SUBAPPLICATION Button_IXA_OR_AX_TO_DataPanel_QXA_BG (* Button (IXA) ODER AX-Eingang auf DataPanel-MI-Ausgang, Hintergrundfarbe Gruen/Weiss, 2 AX-Ausgaenge *)
  (* Standard: 61499-2; Description: Copyright (c) 2026 Meisterschulen am Ostbahnhof This program and the accompanying materials are made available under the terms of the Eclipse Public License 2.0 which is available at https://www.eclipse.org/legal/epl-2.0/ SPDX-License-Identifier: EPL-2.0 *)
  (* Version 1.0, 2026-10-31, Franz Höpfinger, Meisterschulen am Ostbahnhof, Aus Getreidehacke func/Manual/ManFuncTast1 in MyLib::sys verschoben und umbenannt, INIT/INITO/QI/QO ergaenzt, Output und u8SAMember als Parameter. *)
  PACKAGE MyLib::sys;
  IMPORT isobus::UT::Q::const::IDs::ID_NULL;
  IMPORT DataPanel::io::MI::DQ::DataPanel_MI_DO_S;
  IMPORT DataPanel::io::MI::DQ::DataPanel_MI_DO;
  IMPORT DataPanel::io::MI::const::MI;
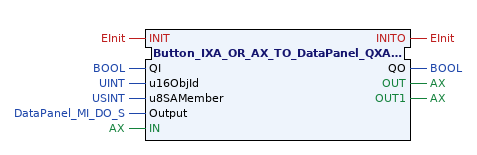
  EVENT_INPUT
    INIT : EInit; (* Initialization Request *)
  END_EVENT
  EVENT_OUTPUT
    INITO : EInit; (* Initialization Confirm *)
  END_EVENT
  VAR_INPUT
    QI : BOOL := TRUE; (* Quality Input - TRUE to enable service *)
    u16ObjId : UINT := ID_NULL; (* Object ID Button *)
    u8SAMember : USINT := MI::MI_00; (* DataPanel-MI-Modul (Source Address) *)
    Output : DataPanel::io::MI::DQ::DataPanel_MI_DO_S := DataPanel_MI_DO::Invalid; (* DataPanel-MI-Ausgang *)
  END_VAR
  VAR_OUTPUT
    QO : BOOL; (* Quality Output - TRUE if service executed successfully *)
  END_VAR
  SOCKETS
    IN : adapter::types::unidirectional::AX; (* zusaetzlicher Eingang, ODER mit Button *)
  END_SOCKETS
  PLUGS
    OUT : adapter::types::unidirectional::AX; (* Button ODER IN *)
    OUT1 : adapter::types::unidirectional::AX; (* Button ODER IN (2. Abgriff) *)
  END_PLUGS
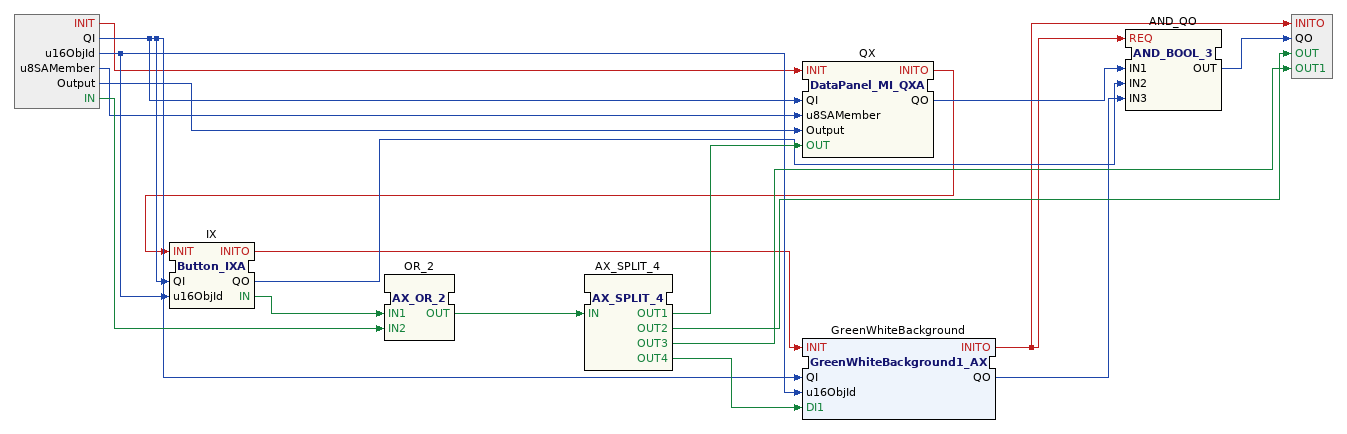
  FBS
    QX : DataPanel::io::MI::DQ::DataPanel_MI_QXA;
    IX : isobus::UT::io::Button::Button_IXA;
    OR_2 : adapter::booleanOperators::AX_OR_2;
    AX_SPLIT_4 : adapter::events::unidirectional::AX_SPLIT_4;
    AND_QO : iec61131::booleanOperators::AND_BOOL_3;
  END_FBS
  SUBAPPS
    GreenWhiteBackground : MyLib::sys::GreenWhiteBackground1_AX;
  END_SUBAPPS
  EVENT_CONNECTIONS
    INIT TO QX.INIT;
    QX.INITO TO IX.INIT;
    IX.INITO TO GreenWhiteBackground.INIT;
    GreenWhiteBackground.INITO TO INITO;
    GreenWhiteBackground.INITO TO AND_QO.REQ;
  END_CONNECTIONS
  DATA_CONNECTIONS
    QI TO QX.QI;
    QI TO IX.QI;
    QI TO GreenWhiteBackground.QI;
    u16ObjId TO IX.u16ObjId;
    u16ObjId TO GreenWhiteBackground.u16ObjId;
    u8SAMember TO QX.u8SAMember;
    Output TO QX.Output;
    QX.QO TO AND_QO.IN1;
    IX.QO TO AND_QO.IN2;
    GreenWhiteBackground.QO TO AND_QO.IN3;
    AND_QO.OUT TO QO;
  END_CONNECTIONS
  ADAPTER_CONNECTIONS
    IX.IN TO OR_2.IN1;
    IN TO OR_2.IN2;
    OR_2.OUT TO AX_SPLIT_4.IN;
    AX_SPLIT_4.OUT1 TO QX.OUT;
    AX_SPLIT_4.OUT2 TO OUT;
    AX_SPLIT_4.OUT3 TO OUT1;
    AX_SPLIT_4.OUT4 TO GreenWhiteBackground.DI1;
  END_CONNECTIONS
END_SUBAPPLICATION
